DATA_BLOCK "FRK_ProductionScratch"
{ S7_Optimized_Access := 'TRUE' }
VERSION : 0.1
NON_RETAIN
VAR
    Calendar {ExternalAccessible := 'False'; ExternalVisible := 'False'; ExternalWritable := 'False'} : "ST_ShiftCalendarV3";
END_VAR
BEGIN
END_DATA_BLOCK
